(* IEC 61131-3 sources: model-first-plc-agent-ai/results/T2-W-07, 2 files *)

(* ---- a1_code.st ---- *)
FUNCTION_BLOCK FB_TimedFilling
VAR_INPUT
    start : BOOL;
    stop : BOOL;
    LSH : BOOL;
    LSHH : BOOL;
    TimerDuration : TIME;
END_VAR
VAR_OUTPUT
    fill_valve : BOOL;
    discharge_valve : BOOL;
END_VAR
VAR
    x0 : BOOL := TRUE;
    x1 : BOOL := FALSE;
    timer_done : BOOL := FALSE;
    FillingTimer : TON;
END_VAR

FillingTimer(IN := x1, PT := TimerDuration);
timer_done := FillingTimer.Q;

IF x1 THEN
    IF stop OR LSHH OR timer_done THEN
        x1 := FALSE;
        x0 := TRUE;

        FillingTimer(IN := FALSE, PT := TimerDuration);
        timer_done := FALSE;
    END_IF;
ELSIF x0 THEN
    IF start AND NOT stop AND NOT LSHH THEN
        x0 := FALSE;
        x1 := TRUE;

        FillingTimer(IN := TRUE, PT := TimerDuration);
        timer_done := FALSE;
    END_IF;
END_IF;

fill_valve := x1;
discharge_valve := FALSE;

END_FUNCTION_BLOCK

PROGRAM Main
VAR
    StartCommand AT %IX100.0 : BOOL;
    StopCommand AT %IX100.1 : BOOL;
    LSH AT %IX100.2 : BOOL;
    LSHH AT %IX100.3 : BOOL;

    FillValve AT %QX100.0 : BOOL;
    DischargeValve AT %QX100.1 : BOOL;
END_VAR
VAR
    (* Configurable filling duration; adjust for the application. *)
    TimerDuration : TIME := T#10s;
    StartEdge : R_TRIG;
    FillingControl : FB_TimedFilling;
END_VAR

StartEdge(CLK := StartCommand);

FillingControl(
    start := StartEdge.Q,
    stop := StopCommand,
    LSH := LSH,
    LSHH := LSHH,
    TimerDuration := TimerDuration
);

FillValve := FillingControl.fill_valve;
DischargeValve := FillingControl.discharge_valve;

END_PROGRAM

(* ---- a2_code.st ---- *)
FUNCTION_BLOCK FB_TankFilling
VAR_INPUT
    StartCommand : BOOL;
    StopCommand : BOOL;
    LSH : BOOL;
    LSHH : BOOL;
    TimerDuration : TIME;
END_VAR
VAR_OUTPUT
    fill_valve : BOOL;
    discharge_valve : BOOL;
END_VAR
VAR
    StateIndex : INT := 0;
    StartEdge : R_TRIG;
    FillingTimer : TON;
    start : BOOL;
    stop : BOOL;
    timer_done : BOOL;
END_VAR

StartEdge(CLK := StartCommand);
start := StartEdge.Q;
stop := StopCommand;

IF stop THEN
    StateIndex := 0;
ELSE
    CASE StateIndex OF
        0:
            IF start THEN
                StateIndex := 1;
            END_IF;
        1:
            StateIndex := 1;
    ELSE
        StateIndex := 0;
    END_CASE;
END_IF;

FillingTimer(IN := (StateIndex = 1), PT := TimerDuration);
timer_done := FillingTimer.Q;

IF (StateIndex = 1) AND (stop OR timer_done OR LSHH) THEN
    StateIndex := 0;
    FillingTimer(IN := FALSE, PT := TimerDuration);
    timer_done := FALSE;
END_IF;

fill_valve := (StateIndex = 1) AND NOT stop;
discharge_valve := FALSE;

END_FUNCTION_BLOCK

PROGRAM Main
VAR
    StartCommand AT %IX100.0 : BOOL;
    StopCommand AT %IX100.1 : BOOL;
    LSH AT %IX100.2 : BOOL;
    LSHH AT %IX100.3 : BOOL;
    FillValve AT %QX100.0 : BOOL;
    DischargeValve AT %QX100.1 : BOOL;
END_VAR
VAR
    TimerDuration : TIME := T#10s;
    TankController : FB_TankFilling;
END_VAR

TankController(
    StartCommand := StartCommand,
    StopCommand := StopCommand,
    LSH := LSH,
    LSHH := LSHH,
    TimerDuration := TimerDuration
);

FillValve := TankController.fill_valve;
DischargeValve := TankController.discharge_valve;

END_PROGRAM
